(* IEC 61131-3 sources: sis-interlock-demo/tests/POUs/Suites/FB_SisEventLog_Test, 7 files *)

(* ---- ClearKeepsSeq.method.decl.st ---- *)
// Clear: записей 0, номер последнего события сохраняется, следующее событие — следующий номер
METHOD PRIVATE ClearKeepsSeq
VAR
    fbLog : FB_SisEventLog;   // журнал
    stEv  : ST_SisEvent;      // событие
END_VAR

(* ---- GetEventBeyondCountEmpty.method.decl.st ---- *)
// GetEvent(uiBack >= Count) — пустая запись: все поля 0
METHOD PRIVATE GetEventBeyondCountEmpty
VAR
    fbLog : FB_SisEventLog;   // журнал
    stEv  : ST_SisEvent;      // событие
END_VAR

(* ---- RingOverwritesOldest.method.decl.st ---- *)
// 70 событий в кольцо на 64: Count = 64, последнее — номер 70, самое старое — номер 7
METHOD PRIVATE RingOverwritesOldest
VAR
    fbLog  : FB_SisEventLog;   // журнал
    stEv   : ST_SisEvent;      // событие
    uiI    : UINT;             // счётчик
    xAdded : BOOL;             // результат записи
    xAll   : BOOL := TRUE;     // все записи приняты
END_VAR

(* ---- RingOverwritesOldest.method.impl.st ---- *)
coUnit.TEST('Log_Ring_OverwritesOldest');
stEv.eKind := E_SisEventKind.CauseDemand;
FOR uiI := 1 TO 70 DO
    stEv.uiCause := uiI;
    xAdded := fbLog.AddEvent(stEvent := stEv);
    xAll := xAll AND xAdded;
END_FOR
AssertTrue(Condition := xAll, Message := 'AddEvent always TRUE');
AssertEquals_UINT(Expected := 64, Actual := fbLog.Count, Message := 'ring full: 64');
AssertEquals_UDINT(Expected := 70, Actual := fbLog.LastSeq, Message := 'last seq 70');
stEv := fbLog.GetEvent(uiBack := 0);
AssertEquals_UDINT(Expected := 70, Actual := stEv.udiSeq, Message := 'newest: seq 70');
AssertEquals_UINT(Expected := 70, Actual := stEv.uiCause, Message := 'newest: cause 70');
stEv := fbLog.GetEvent(uiBack := 63);
AssertEquals_UDINT(Expected := 7, Actual := stEv.udiSeq, Message := 'oldest kept: seq 7');
AssertEquals_UINT(Expected := 7, Actual := stEv.uiCause, Message := 'oldest kept: cause 7');
coUnit.TEST_FINISHED();

(* ---- SeqIncrementsAndWraps.method.decl.st ---- *)
// Номер события растёт на 1; после 16#FFFFFFFF — снова 1 (0 не выдаётся)
METHOD PRIVATE SeqIncrementsAndWraps
VAR
    fbLog : FB_SisTestLog;    // журнал с установкой номера
    stEv  : ST_SisEvent;      // событие
END_VAR

(* ---- SizeOfEventIs24.method.decl.st ---- *)
// Запись журнала — 24 байта без выравнивающих пропусков (раздел 4.2)
METHOD PRIVATE SizeOfEventIs24
VAR
    stEv : ST_SisEvent;   // запись
END_VAR

(* ---- ViaInterfaceKeepsFields.method.decl.st ---- *)
// Запись через I_SisEventSink: все поля, кроме номера, сохраняются как есть
METHOD PRIVATE ViaInterfaceKeepsFields
VAR
    fbLog  : FB_SisEventLog;   // журнал
    itfLog : I_SisEventSink;   // журнал как приёмник
    stEv   : ST_SisEvent;      // событие
    stGot  : ST_SisEvent;      // прочитанное событие
    xAdded : BOOL;             // результат записи
END_VAR
